(*!
<summary>Formats a failed typed predicate and reports it with the chain message.</summary>
<description>
Does not change operands or chain state. The receiver retains its first failure. Reporting exceptions
propagate to the enclosing test callback handler; an unprepared receiver is a configuration error.
</description>
<param name="expected">Typed expected operand used only for this diagnostic.</param>
<param name="expectation">Prefix identifying the failed predicate.</param>
*)
METHOD PRIVATE failComparison
VAR_INPUT
	expected : SINT;
	expectation : WSTRING(40);
END_VAR
VAR
	actualText : WSTRING(255);
	expectedText : WSTRING(255);
	diagnostic : TOF_Core.ERROR_MESSAGE;
END_VAR
actualText := TO_WSTRING(_Actual);
expectedText := TO_WSTRING(expected);

diagnostic := TOF_Core.WideStrings.Concat255(
	expectation,
	expectedText,
	", but was: ",
	actualText
);

TestServices.ReportAssertionFailure(
	testCase := _TestCase,
	message := _Message,
	sourceClassName := ClassName,
	defaultMessage := diagnostic
);
END_METHOD

END_FUNCTION_BLOCK

// ---- Assertions/TypedContexts/IntAssertionContext.TcPOU
(*
SPDX-FileCopyrightText: © 2026 Oleksandr Tiutyk <trofimich@gmail.com>
SPDX-License-Identifier: MIT
License: https://opensource.org/license/mit
*)

(*!
<summary>Provides fluent assertions on a copied INT value.</summary>
<description>
Copies actual into persistent instance storage before the entry method returns; literals and expression
results therefore remain valid throughout the immediate chain. Owns no heap allocation or pointed-to resource.
The message prefixes every failure until the next preparation. Finish one chain before starting another on
the owning Assertions provider. Use only from the owning test callback on one task, without reentry.
Obtain this context from the owning provider; direct unprepared use is unsupported.
Expected arguments use the declared IEC type; ordinary compiler conversions happen before comparison.
This context does not depend on another assertion context.
Object metadata is available before preparation; inherited equality compares instance identity.
</description>
*)

{attribute 'no_explicit_call' := 'do not call this function block directly'}
FUNCTION_BLOCK IntAssertionContext EXTENDS TOF_Core.Object
VAR_STAT
	{attribute 'hide'}
	_ClassName : STRING := __POUNAME();
END_VAR
VAR
	_Actual : INT;
	_TestCase : ITestCase;
	_Message : WSTRING(255);
END_VAR

(*!
<summary>Provides the implementation class name.</summary>
<description>
Borrowed read-only reference to compiler-initialized storage, valid throughout the instance lifetime.
Do not modify the returned reference; no ownership is transferred.
</description>
*)
{attribute 'monitoring' := 'call'}
PROPERTY ClassName : REFERENCE TO STRING
GET
ClassName REF= _ClassName;
END_GET
END_PROPERTY

(*!
<summary>Asserts that the actual value is strictly greater than expected.</summary>
<description>
Records failure without interrupting the callback; preserves the message for the rest of the chain.
</description>
<param name="expected">Expected value converted by the compiler to INT.</param>
*)
METHOD FINAL IsGreaterThan : REFERENCE TO IntAssertionContext
VAR_INPUT
	expected : INT;
END_VAR
IF _Actual <= expected THEN
	failComparison(
		expected := expected,
		expectation := "Expected value > "
	);
END_IF

IsGreaterThan REF= THIS^;
END_METHOD

(*!
<summary>Asserts that the actual value meets the inclusive lower boundary.</summary>
<description>
Records failure without interrupting the callback; preserves the message for the rest of the chain.
</description>
<param name="expected">Expected value converted by the compiler to INT.</param>
*)
METHOD FINAL IsGreaterThanOrEquals : REFERENCE TO IntAssertionContext
VAR_INPUT
	expected : INT;
END_VAR
IF _Actual < expected THEN
	failComparison(
		expected := expected,
		expectation := "Expected value >= "
	);
END_IF

IsGreaterThanOrEquals REF= THIS^;
END_METHOD

(*!
<summary>Asserts that the actual value is strictly less than expected.</summary>
<description>
Records failure without interrupting the callback; preserves the message for the rest of the chain.
</description>
<param name="expected">Expected value converted by the compiler to INT.</param>
*)
METHOD FINAL IsLessThan : REFERENCE TO IntAssertionContext
VAR_INPUT
	expected : INT;
END_VAR
IF _Actual >= expected THEN
	failComparison(
		expected := expected,
		expectation := "Expected value < "
	);
END_IF

IsLessThan REF= THIS^;
END_METHOD

(*!
<summary>Asserts that the actual value meets the inclusive upper boundary.</summary>
<description>
Records failure without interrupting the callback; preserves the message for the rest of the chain.
</description>
<param name="expected">Expected value converted by the compiler to INT.</param>
*)
METHOD FINAL IsLessThanOrEquals : REFERENCE TO IntAssertionContext
VAR_INPUT
	expected : INT;
END_VAR
IF _Actual > expected THEN
	failComparison(
		expected := expected,
		expectation := "Expected value <= "
	);
END_IF

IsLessThanOrEquals REF= THIS^;
END_METHOD

(*!
<summary>Provides the library namespace.</summary>
<description>
Borrowed read-only reference to the compiler-initialized namespace, valid throughout the instance lifetime.
Do not modify the returned reference; no ownership is transferred.
</description>
*)
{attribute 'monitoring' := 'call'}
PROPERTY NamespaceName : REFERENCE TO STRING
GET
NamespaceName REF= CurrentNamespace.Name;
END_GET
END_PROPERTY

(*!
<summary>Asserts inequality with the expected value.</summary>
<description>
Records failure without interrupting the callback; preserves the message for the rest of the chain.
</description>
<param name="expected">Expected value converted by the compiler to INT.</param>
*)
METHOD FINAL NotToBe : REFERENCE TO IntAssertionContext
VAR_INPUT
	expected : INT;
END_VAR
IF _Actual = expected THEN
	failComparison(
		expected := expected,
		expectation := "Expected value not to be: "
	);
END_IF

NotToBe REF= THIS^;
END_METHOD

(*!
<summary>Copies the actual operand and replaces the chain-wide message.</summary>
<description>
Called by the owning Assertions provider after it verifies the running test case.
No pointer to this method's input storage is retained. The receiver is borrowed until the next preparation;
the owning provider keeps it alive throughout the immediate chain.
</description>
<param name="actual">Value copied into this context.</param>
<param name="testCase">Borrowed failure receiver for the immediate chain.</param>
<param name="message">Copied diagnostic prefix, including empty to clear the previous prefix.</param>
*)
METHOD INTERNAL FINAL Prepare
VAR_INPUT
	actual : INT;
	testCase : ITestCase;
	message : WSTRING(255);
END_VAR
_Actual := actual;
_TestCase := testCase;
_Message := message;
END_METHOD

(*!
<summary>Reports the byte size of this concrete instance.</summary>
<description>
Includes inline fields and nested instances, but excludes separately allocated payloads.
Obtaining the size does not transfer ownership or validate an arbitrary address.
</description>
*)
{attribute 'monitoring' := 'call'}
PROPERTY SelfSize : ULINT
GET
SelfSize := XSIZEOF(THIS^);
END_GET
END_PROPERTY

(*!
<summary>Asserts equality with the expected value.</summary>
<description>
Records failure without interrupting the callback; preserves the message for the rest of the chain.
</description>
<param name="expected">Expected value converted by the compiler to INT.</param>
*)
METHOD FINAL ToBe : REFERENCE TO IntAssertionContext
VAR_INPUT
	expected : INT;
END_VAR
IF _Actual <> expected THEN
	failComparison(
		expected := expected,
		expectation := "Expected: "
	);
END_IF

ToBe REF= THIS^;
END_METHOD

(*!
<summary>Formats a failed typed predicate and reports it with the chain message.</summary>
<description>
Does not change operands or chain state. The receiver retains its first failure. Reporting exceptions
propagate to the enclosing test callback handler; an unprepared receiver is a configuration error.
</description>
<param name="expected">Typed expected operand used only for this diagnostic.</param>
<param name="expectation">Prefix identifying the failed predicate.</param>
*)
METHOD PRIVATE failComparison
VAR_INPUT
	expected : INT;
	expectation : WSTRING(40);
END_VAR
VAR
	actualText : WSTRING(255);
	expectedText : WSTRING(255);
	diagnostic : TOF_Core.ERROR_MESSAGE;
END_VAR
actualText := TO_WSTRING(_Actual);
expectedText := TO_WSTRING(expected);

diagnostic := TOF_Core.WideStrings.Concat255(
	expectation,
	expectedText,
	", but was: ",
	actualText
);

TestServices.ReportAssertionFailure(
	testCase := _TestCase,
	message := _Message,
	sourceClassName := ClassName,
	defaultMessage := diagnostic
);
END_METHOD

END_FUNCTION_BLOCK

// ---- Assertions/TypedContexts/DIntAssertionContext.TcPOU
(*
SPDX-FileCopyrightText: © 2026 Oleksandr Tiutyk <trofimich@gmail.com>
SPDX-License-Identifier: MIT
License: https://opensource.org/license/mit
*)

(*!
<summary>Provides fluent assertions on a copied DINT value.</summary>
<description>
Copies actual into persistent instance storage before the entry method returns; literals and expression
results therefore remain valid throughout the immediate chain. Owns no heap allocation or pointed-to resource.
The message prefixes every failure until the next preparation. Finish one chain before starting another on
the owning Assertions provider. Use only from the owning test callback on one task, without reentry.
Obtain this context from the owning provider; direct unprepared use is unsupported.
Expected arguments use the declared IEC type; ordinary compiler conversions happen before comparison.
This context does not depend on another assertion context.
Object metadata is available before preparation; inherited equality compares instance identity.
</description>
*)

{attribute 'no_explicit_call' := 'do not call this function block directly'}
FUNCTION_BLOCK DIntAssertionContext EXTENDS TOF_Core.Object
VAR_STAT
	{attribute 'hide'}
	_ClassName : STRING := __POUNAME();
END_VAR
VAR
	_Actual : DINT;
	_TestCase : ITestCase;
	_Message : WSTRING(255);
END_VAR

(*!
<summary>Provides the implementation class name.</summary>
<description>
Borrowed read-only reference to compiler-initialized storage, valid throughout the instance lifetime.
Do not modify the returned reference; no ownership is transferred.
</description>
*)
{attribute 'monitoring' := 'call'}
PROPERTY ClassName : REFERENCE TO STRING
GET
ClassName REF= _ClassName;
END_GET
END_PROPERTY

(*!
<summary>Asserts that the actual value is strictly greater than expected.</summary>
<description>
Records failure without interrupting the callback; preserves the message for the rest of the chain.
</description>
<param name="expected">Expected value converted by the compiler to DINT.</param>
*)
METHOD FINAL IsGreaterThan : REFERENCE TO DIntAssertionContext
VAR_INPUT
	expected : DINT;
END_VAR
IF _Actual <= expected THEN
	failComparison(
		expected := expected,
		expectation := "Expected value > "
	);
END_IF

IsGreaterThan REF= THIS^;
END_METHOD

(*!
<summary>Asserts that the actual value meets the inclusive lower boundary.</summary>
<description>
Records failure without interrupting the callback; preserves the message for the rest of the chain.
</description>
<param name="expected">Expected value converted by the compiler to DINT.</param>
*)
METHOD FINAL IsGreaterThanOrEquals : REFERENCE TO DIntAssertionContext
VAR_INPUT
	expected : DINT;
END_VAR
IF _Actual < expected THEN
	failComparison(
		expected := expected,
		expectation := "Expected value >= "
	);
END_IF

IsGreaterThanOrEquals REF= THIS^;
END_METHOD

(*!
<summary>Asserts that the actual value is strictly less than expected.</summary>
<description>
Records failure without interrupting the callback; preserves the message for the rest of the chain.
</description>
<param name="expected">Expected value converted by the compiler to DINT.</param>
*)
METHOD FINAL IsLessThan : REFERENCE TO DIntAssertionContext
VAR_INPUT
	expected : DINT;
END_VAR
IF _Actual >= expected THEN
	failComparison(
		expected := expected,
		expectation := "Expected value < "
	);
END_IF

IsLessThan REF= THIS^;
END_METHOD

(*!
<summary>Asserts that the actual value meets the inclusive upper boundary.</summary>
<description>
Records failure without interrupting the callback; preserves the message for the rest of the chain.
</description>
<param name="expected">Expected value converted by the compiler to DINT.</param>
*)
METHOD FINAL IsLessThanOrEquals : REFERENCE TO DIntAssertionContext
VAR_INPUT
	expected : DINT;
END_VAR
IF _Actual > expected THEN
	failComparison(
		expected := expected,
		expectation := "Expected value <= "
	);
END_IF

IsLessThanOrEquals REF= THIS^;
END_METHOD

(*!
<summary>Provides the library namespace.</summary>
<description>
Borrowed read-only reference to the compiler-initialized namespace, valid throughout the instance lifetime.
Do not modify the returned reference; no ownership is transferred.
</description>
*)
{attribute 'monitoring' := 'call'}
PROPERTY NamespaceName : REFERENCE TO STRING
GET
NamespaceName REF= CurrentNamespace.Name;
END_GET
END_PROPERTY

(*!
<summary>Asserts inequality with the expected value.</summary>
<description>
Records failure without interrupting the callback; preserves the message for the rest of the chain.
</description>
<param name="expected">Expected value converted by the compiler to DINT.</param>
*)
METHOD FINAL NotToBe : REFERENCE TO DIntAssertionContext
VAR_INPUT
	expected : DINT;
END_VAR
IF _Actual = expected THEN
	failComparison(
		expected := expected,
		expectation := "Expected value not to be: "
	);
END_IF

NotToBe REF= THIS^;
END_METHOD

(*!
<summary>Copies the actual operand and replaces the chain-wide message.</summary>
<description>
Called by the owning Assertions provider after it verifies the running test case.
No pointer to this method's input storage is retained. The receiver is borrowed until the next preparation;
the owning provider keeps it alive throughout the immediate chain.
</description>
<param name="actual">Value copied into this context.</param>
<param name="testCase">Borrowed failure receiver for the immediate chain.</param>
<param name="message">Copied diagnostic prefix, including empty to clear the previous prefix.</param>
*)
METHOD INTERNAL FINAL Prepare
VAR_INPUT
	actual : DINT;
	testCase : ITestCase;
	message : WSTRING(255);
END_VAR
_Actual := actual;
_TestCase := testCase;
_Message := message;
END_METHOD

(*!
<summary>Reports the byte size of this concrete instance.</summary>
<description>
Includes inline fields and nested instances, but excludes separately allocated payloads.
Obtaining the size does not transfer ownership or validate an arbitrary address.
</description>
*)
{attribute 'monitoring' := 'call'}
PROPERTY SelfSize : ULINT
GET
SelfSize := XSIZEOF(THIS^);
END_GET
END_PROPERTY

(*!
<summary>Asserts equality with the expected value.</summary>
<description>
Records failure without interrupting the callback; preserves the message for the rest of the chain.
</description>
<param name="expected">Expected value converted by the compiler to DINT.</param>
*)
METHOD FINAL ToBe : REFERENCE TO DIntAssertionContext
VAR_INPUT
	expected : DINT;
END_VAR
IF _Actual <> expected THEN
	failComparison(
		expected := expected,
		expectation := "Expected: "
	);
END_IF

ToBe REF= THIS^;
END_METHOD

(*!
<summary>Formats a failed typed predicate and reports it with the chain message.</summary>
<description>
Does not change operands or chain state. The receiver retains its first failure. Reporting exceptions
propagate to the enclosing test callback handler; an unprepared receiver is a configuration error.
</description>
<param name="expected">Typed expected operand used only for this diagnostic.</param>
<param name="expectation">Prefix identifying the failed predicate.</param>
*)
METHOD PRIVATE failComparison
VAR_INPUT
	expected : DINT;
	expectation : WSTRING(40);
END_VAR
VAR
	actualText : WSTRING(255);
	expectedText : WSTRING(255);
	diagnostic : TOF_Core.ERROR_MESSAGE;
END_VAR
actualText := TO_WSTRING(_Actual);
expectedText := TO_WSTRING(expected);

diagnostic := TOF_Core.WideStrings.Concat255(
	expectation,
	expectedText,
	", but was: ",
	actualText
);

TestServices.ReportAssertionFailure(
	testCase := _TestCase,
	message := _Message,
	sourceClassName := ClassName,
	defaultMessage := diagnostic
);
END_METHOD

END_FUNCTION_BLOCK

// ---- Assertions/TypedContexts/LIntAssertionContext.TcPOU
(*
SPDX-FileCopyrightText: © 2026 Oleksandr Tiutyk <trofimich@gmail.com>
SPDX-License-Identifier: MIT
License: https://opensource.org/license/mit
*)

(*!
<summary>Provides fluent assertions on a copied LINT value.</summary>
<description>
Copies actual into persistent instance storage before the entry method returns; literals and expression
results therefore remain valid throughout the immediate chain. Owns no heap allocation or pointed-to resource.
The message prefixes every failure until the next preparation. Finish one chain before starting another on
the owning Assertions provider. Use only from the owning test callback on one task, without reentry.
Obtain this context from the owning provider; direct unprepared use is unsupported.
Expected arguments use the declared IEC type; ordinary compiler conversions happen before comparison.
This context does not depend on another assertion context.
Object metadata is available before preparation; inherited equality compares instance identity.
</description>
*)

{attribute 'no_explicit_call' := 'do not call this function block directly'}
FUNCTION_BLOCK LIntAssertionContext EXTENDS TOF_Core.Object
VAR_STAT
	{attribute 'hide'}
	_ClassName : STRING := __POUNAME();
END_VAR
VAR
	_Actual : LINT;
	_TestCase : ITestCase;
	_Message : WSTRING(255);
END_VAR

(*!
<summary>Provides the implementation class name.</summary>
<description>
Borrowed read-only reference to compiler-initialized storage, valid throughout the instance lifetime.
Do not modify the returned reference; no ownership is transferred.
</description>
*)
{attribute 'monitoring' := 'call'}
PROPERTY ClassName : REFERENCE TO STRING
GET
ClassName REF= _ClassName;
END_GET
END_PROPERTY

(*!
<summary>Asserts that the actual value is strictly greater than expected.</summary>
<description>
Records failure without interrupting the callback; preserves the message for the rest of the chain.
</description>
<param name="expected">Expected value converted by the compiler to LINT.</param>
*)
METHOD FINAL IsGreaterThan : REFERENCE TO LIntAssertionContext
VAR_INPUT
	expected : LINT;
END_VAR
IF _Actual <= expected THEN
	failComparison(
		expected := expected,
		expectation := "Expected value > "
	);
END_IF

IsGreaterThan REF= THIS^;
END_METHOD

(*!
<summary>Asserts that the actual value meets the inclusive lower boundary.</summary>
<description>
Records failure without interrupting the callback; preserves the message for the rest of the chain.
</description>
<param name="expected">Expected value converted by the compiler to LINT.</param>
*)
METHOD FINAL IsGreaterThanOrEquals : REFERENCE TO LIntAssertionContext
VAR_INPUT
	expected : LINT;
END_VAR
IF _Actual < expected THEN
	failComparison(
		expected := expected,
		expectation := "Expected value >= "
	);
END_IF

IsGreaterThanOrEquals REF= THIS^;
END_METHOD

(*!
<summary>Asserts that the actual value is strictly less than expected.</summary>
<description>
Records failure without interrupting the callback; preserves the message for the rest of the chain.
</description>
<param name="expected">Expected value converted by the compiler to LINT.</param>
*)
METHOD FINAL IsLessThan : REFERENCE TO LIntAssertionContext
VAR_INPUT
	expected : LINT;
END_VAR
IF _Actual >= expected THEN
	failComparison(
		expected := expected,
		expectation := "Expected value < "
	);
END_IF

IsLessThan REF= THIS^;
END_METHOD

(*!
<summary>Asserts that the actual value meets the inclusive upper boundary.</summary>
<description>
Records failure without interrupting the callback; preserves the message for the rest of the chain.
</description>
<param name="expected">Expected value converted by the compiler to LINT.</param>
*)
METHOD FINAL IsLessThanOrEquals : REFERENCE TO LIntAssertionContext
VAR_INPUT
	expected : LINT;
END_VAR
IF _Actual > expected THEN
	failComparison(
		expected := expected,
		expectation := "Expected value <= "
	);
END_IF

IsLessThanOrEquals REF= THIS^;
END_METHOD

(*!
<summary>Provides the library namespace.</summary>
<description>
Borrowed read-only reference to the compiler-initialized namespace, valid throughout the instance lifetime.
Do not modify the returned reference; no ownership is transferred.
</description>
*)
{attribute 'monitoring' := 'call'}
PROPERTY NamespaceName : REFERENCE TO STRING
GET
NamespaceName REF= CurrentNamespace.Name;
END_GET
END_PROPERTY

(*!
<summary>Asserts inequality with the expected value.</summary>
<description>
Records failure without interrupting the callback; preserves the message for the rest of the chain.
</description>
<param name="expected">Expected value converted by the compiler to LINT.</param>
*)
METHOD FINAL NotToBe : REFERENCE TO LIntAssertionContext
VAR_INPUT
	expected : LINT;
END_VAR
IF _Actual = expected THEN
	failComparison(
		expected := expected,
		expectation := "Expected value not to be: "
	);
END_IF

NotToBe REF= THIS^;
END_METHOD

(*!
<summary>Copies the actual operand and replaces the chain-wide message.</summary>
<description>
Called by the owning Assertions provider after it verifies the running test case.
No pointer to this method's input storage is retained. The receiver is borrowed until the next preparation;
the owning provider keeps it alive throughout the immediate chain.
</description>
<param name="actual">Value copied into this context.</param>
<param name="testCase">Borrowed failure receiver for the immediate chain.</param>
<param name="message">Copied diagnostic prefix, including empty to clear the previous prefix.</param>
*)
METHOD INTERNAL FINAL Prepare
VAR_INPUT
	actual : LINT;
	testCase : ITestCase;
	message : WSTRING(255);
END_VAR
_Actual := actual;
_TestCase := testCase;
_Message := message;
END_METHOD

(*!
<summary>Reports the byte size of this concrete instance.</summary>
<description>
Includes inline fields and nested instances, but excludes separately allocated payloads.
Obtaining the size does not transfer ownership or validate an arbitrary address.
</description>
*)
{attribute 'monitoring' := 'call'}
PROPERTY SelfSize : ULINT
GET
SelfSize := XSIZEOF(THIS^);
END_GET
END_PROPERTY

(*!
<summary>Asserts equality with the expected value.</summary>
<description>
Records failure without interrupting the callback; preserves the message for the rest of the chain.
</description>
<param name="expected">Expected value converted by the compiler to LINT.</param>
*)
METHOD FINAL ToBe : REFERENCE TO LIntAssertionContext
VAR_INPUT
	expected : LINT;
END_VAR
IF _Actual <> expected THEN
	failComparison(
		expected := expected,
		expectation := "Expected: "
	);
END_IF

ToBe REF= THIS^;
END_METHOD

(*!
<summary>Formats a failed typed predicate and reports it with the chain message.</summary>
<description>
Does not change operands or chain state. The receiver retains its first failure. Reporting exceptions
propagate to the enclosing test callback handler; an unprepared receiver is a configuration error.
</description>
<param name="expected">Typed expected operand used only for this diagnostic.</param>
<param name="expectation">Prefix identifying the failed predicate.</param>
*)
METHOD PRIVATE failComparison
VAR_INPUT
	expected : LINT;
	expectation : WSTRING(40);
END_VAR
VAR
	actualText : WSTRING(255);
	expectedText : WSTRING(255);
	diagnostic : TOF_Core.ERROR_MESSAGE;
END_VAR
actualText := TO_WSTRING(_Actual);
expectedText := TO_WSTRING(expected);

diagnostic := TOF_Core.WideStrings.Concat255(
	expectation,
	expectedText,
	", but was: ",
	actualText
);

TestServices.ReportAssertionFailure(
	testCase := _TestCase,
	message := _Message,
	sourceClassName := ClassName,
	defaultMessage := diagnostic
);
END_METHOD

END_FUNCTION_BLOCK

// ---- Assertions/TypedContexts/USIntAssertionContext.TcPOU
(*
SPDX-FileCopyrightText: © 2026 Oleksandr Tiutyk <trofimich@gmail.com>
SPDX-License-Identifier: MIT
License: https://opensource.org/license/mit
*)

(*!
<summary>Provides fluent assertions on a copied USINT value.</summary>
<description>
Copies actual into persistent instance storage before the entry method returns; literals and expression
results therefore remain valid throughout the immediate chain. Owns no heap allocation or pointed-to resource.
The message prefixes every failure until the next preparation. Finish one chain before starting another on
the owning Assertions provider. Use only from the owning test callback on one task, without reentry.
Obtain this context from the owning provider; direct unprepared use is unsupported.
Expected arguments use the declared IEC type; ordinary compiler conversions happen before comparison.
This context does not depend on another assertion context.
Object metadata is available before preparation; inherited equality compares instance identity.
</description>
*)

{attribute 'no_explicit_call' := 'do not call this function block directly'}
FUNCTION_BLOCK USIntAssertionContext EXTENDS TOF_Core.Object
VAR_STAT
	{attribute 'hide'}
	_ClassName : STRING := __POUNAME();
END_VAR
VAR
	_Actual : USINT;
	_TestCase : ITestCase;
	_Message : WSTRING(255);
END_VAR

(*!
<summary>Provides the implementation class name.</summary>
<description>
Borrowed read-only reference to compiler-initialized storage, valid throughout the instance lifetime.
Do not modify the returned reference; no ownership is transferred.
</description>
*)
{attribute 'monitoring' := 'call'}
PROPERTY ClassName : REFERENCE TO STRING
GET
ClassName REF= _ClassName;
END_GET
END_PROPERTY

(*!
<summary>Asserts that the actual value is strictly greater than expected.</summary>
<description>
Records failure without interrupting the callback; preserves the message for the rest of the chain.
</description>
<param name="expected">Expected value converted by the compiler to USINT.</param>
*)
METHOD FINAL IsGreaterThan : REFERENCE TO USIntAssertionContext
VAR_INPUT
	expected : USINT;
END_VAR
IF _Actual <= expected THEN
	failComparison(
		expected := expected,
		expectation := "Expected value > "
	);
END_IF

IsGreaterThan REF= THIS^;
END_METHOD

(*!
<summary>Asserts that the actual value meets the inclusive lower boundary.</summary>
<description>
Records failure without interrupting the callback; preserves the message for the rest of the chain.
</description>
<param name="expected">Expected value converted by the compiler to USINT.</param>
*)
METHOD FINAL IsGreaterThanOrEquals : REFERENCE TO USIntAssertionContext
VAR_INPUT
	expected : USINT;
END_VAR
IF _Actual < expected THEN
	failComparison(
		expected := expected,
		expectation := "Expected value >= "
	);
END_IF

IsGreaterThanOrEquals REF= THIS^;
END_METHOD

(*!
<summary>Asserts that the actual value is strictly less than expected.</summary>
<description>
Records failure without interrupting the callback; preserves the message for the rest of the chain.
</description>
<param name="expected">Expected value converted by the compiler to USINT.</param>
*)
METHOD FINAL IsLessThan : REFERENCE TO USIntAssertionContext
VAR_INPUT
	expected : USINT;
END_VAR
IF _Actual >= expected THEN
	failComparison(
		expected := expected,
		expectation := "Expected value < "
	);
END_IF

IsLessThan REF= THIS^;
END_METHOD

(*!
<summary>Asserts that the actual value meets the inclusive upper boundary.</summary>
<description>
Records failure without interrupting the callback; preserves the message for the rest of the chain.
</description>
<param name="expected">Expected value converted by the compiler to USINT.</param>
*)
METHOD FINAL IsLessThanOrEquals : REFERENCE TO USIntAssertionContext
VAR_INPUT
	expected : USINT;
END_VAR
IF _Actual > expected THEN
	failComparison(
		expected := expected,
		expectation := "Expected value <= "
	);
END_IF

IsLessThanOrEquals REF= THIS^;
END_METHOD

(*!
<summary>Provides the library namespace.</summary>
<description>
Borrowed read-only reference to the compiler-initialized namespace, valid throughout the instance lifetime.
Do not modify the returned reference; no ownership is transferred.
</description>
*)
{attribute 'monitoring' := 'call'}
PROPERTY NamespaceName : REFERENCE TO STRING
GET
NamespaceName REF= CurrentNamespace.Name;
END_GET
END_PROPERTY

(*!
<summary>Asserts inequality with the expected value.</summary>
<description>
Records failure without interrupting the callback; preserves the message for the rest of the chain.
</description>
<param name="expected">Expected value converted by the compiler to USINT.</param>
*)
METHOD FINAL NotToBe : REFERENCE TO USIntAssertionContext
VAR_INPUT
	expected : USINT;
END_VAR
IF _Actual = expected THEN
	failComparison(
		expected := expected,
		expectation := "Expected value not to be: "
	);
END_IF

NotToBe REF= THIS^;
END_METHOD

(*!
<summary>Copies the actual operand and replaces the chain-wide message.</summary>
<description>
Called by the owning Assertions provider after it verifies the running test case.
No pointer to this method's input storage is retained. The receiver is borrowed until the next preparation;
the owning provider keeps it alive throughout the immediate chain.
</description>
<param name="actual">Value copied into this context.</param>
<param name="testCase">Borrowed failure receiver for the immediate chain.</param>
<param name="message">Copied diagnostic prefix, including empty to clear the previous prefix.</param>
*)
METHOD INTERNAL FINAL Prepare
VAR_INPUT
	actual : USINT;
	testCase : ITestCase;
	message : WSTRING(255);
END_VAR
_Actual := actual;
_TestCase := testCase;
_Message := message;
END_METHOD

(*!
<summary>Reports the byte size of this concrete instance.</summary>
<description>
Includes inline fields and nested instances, but excludes separately allocated payloads.
Obtaining the size does not transfer ownership or validate an arbitrary address.
</description>
*)
{attribute 'monitoring' := 'call'}
PROPERTY SelfSize : ULINT
GET
SelfSize := XSIZEOF(THIS^);
END_GET
END_PROPERTY

(*!
<summary>Asserts equality with the expected value.</summary>
<description>
Records failure without interrupting the callback; preserves the message for the rest of the chain.
</description>
<param name="expected">Expected value converted by the compiler to USINT.</param>
*)
METHOD FINAL ToBe : REFERENCE TO USIntAssertionContext
VAR_INPUT
	expected : USINT;
END_VAR
IF _Actual <> expected THEN
	failComparison(
		expected := expected,
		expectation := "Expected: "
	);
END_IF

ToBe REF= THIS^;
END_METHOD

(*!
<summary>Formats a failed typed predicate and reports it with the chain message.</summary>
<description>
Does not change operands or chain state. The receiver retains its first failure. Reporting exceptions
propagate to the enclosing test callback handler; an unprepared receiver is a configuration error.
</description>
<param name="expected">Typed expected operand used only for this diagnostic.</param>
<param name="expectation">Prefix identifying the failed predicate.</param>
*)
METHOD PRIVATE failComparison
VAR_INPUT
	expected : USINT;
	expectation : WSTRING(40);
END_VAR
VAR
	actualText : WSTRING(255);
	expectedText : WSTRING(255);
	diagnostic : TOF_Core.ERROR_MESSAGE;
END_VAR
actualText := TO_WSTRING(_Actual);
expectedText := TO_WSTRING(expected);

diagnostic := TOF_Core.WideStrings.Concat255(
	expectation,
	expectedText,
	", but was: ",
	actualText
);

TestServices.ReportAssertionFailure(
	testCase := _TestCase,
	message := _Message,
	sourceClassName := ClassName,
	defaultMessage := diagnostic
);
END_METHOD

END_FUNCTION_BLOCK

// ---- Assertions/TypedContexts/UIntAssertionContext.TcPOU
(*
SPDX-FileCopyrightText: © 2026 Oleksandr Tiutyk <trofimich@gmail.com>
SPDX-License-Identifier: MIT
License: https://opensource.org/license/mit
*)

(*!
<summary>Provides fluent assertions on a copied UINT value.</summary>
<description>
Copies actual into persistent instance storage before the entry method returns; literals and expression
results therefore remain valid throughout the immediate chain. Owns no heap allocation or pointed-to resource.
The message prefixes every failure until the next preparation. Finish one chain before starting another on
the owning Assertions provider. Use only from the owning test callback on one task, without reentry.
Obtain this context from the owning provider; direct unprepared use is unsupported.
Expected arguments use the declared IEC type; ordinary compiler conversions happen before comparison.
This context does not depend on another assertion context.
Object metadata is available before preparation; inherited equality compares instance identity.
</description>
*)

{attribute 'no_explicit_call' := 'do not call this function block directly'}
FUNCTION_BLOCK UIntAssertionContext EXTENDS TOF_Core.Object
VAR_STAT
	{attribute 'hide'}
	_ClassName : STRING := __POUNAME();
END_VAR
VAR
	_Actual : UINT;
	_TestCase : ITestCase;
	_Message : WSTRING(255);
END_VAR

(*!
<summary>Provides the implementation class name.</summary>
<description>
Borrowed read-only reference to compiler-initialized storage, valid throughout the instance lifetime.
Do not modify the returned reference; no ownership is transferred.
</description>
*)
{attribute 'monitoring' := 'call'}
PROPERTY ClassName : REFERENCE TO STRING
GET
ClassName REF= _ClassName;
END_GET
END_PROPERTY

(*!
<summary>Asserts that the actual value is strictly greater than expected.</summary>
<description>
Records failure without interrupting the callback; preserves the message for the rest of the chain.
</description>
<param name="expected">Expected value converted by the compiler to UINT.</param>
*)
METHOD FINAL IsGreaterThan : REFERENCE TO UIntAssertionContext
VAR_INPUT
	expected : UINT;
END_VAR
IF _Actual <= expected THEN
	failComparison(
		expected := expected,
		expectation := "Expected value > "
	);
END_IF

IsGreaterThan REF= THIS^;
END_METHOD

(*!
<summary>Asserts that the actual value meets the inclusive lower boundary.</summary>
<description>
Records failure without interrupting the callback; preserves the message for the rest of the chain.
</description>
<param name="expected">Expected value converted by the compiler to UINT.</param>
*)
METHOD FINAL IsGreaterThanOrEquals : REFERENCE TO UIntAssertionContext
VAR_INPUT
	expected : UINT;
END_VAR
IF _Actual < expected THEN
	failComparison(
		expected := expected,
		expectation := "Expected value >= "
	);
END_IF

IsGreaterThanOrEquals REF= THIS^;
END_METHOD

(*!
<summary>Asserts that the actual value is strictly less than expected.</summary>
<description>
Records failure without interrupting the callback; preserves the message for the rest of the chain.
</description>
<param name="expected">Expected value converted by the compiler to UINT.</param>
*)
METHOD FINAL IsLessThan : REFERENCE TO UIntAssertionContext
VAR_INPUT
	expected : UINT;
END_VAR
IF _Actual >= expected THEN
	failComparison(
		expected := expected,
		expectation := "Expected value < "
	);
END_IF

IsLessThan REF= THIS^;
END_METHOD

(*!
<summary>Asserts that the actual value meets the inclusive upper boundary.</summary>
<description>
Records failure without interrupting the callback; preserves the message for the rest of the chain.
</description>
<param name="expected">Expected value converted by the compiler to UINT.</param>
*)
METHOD FINAL IsLessThanOrEquals : REFERENCE TO UIntAssertionContext
VAR_INPUT
	expected : UINT;
END_VAR
IF _Actual > expected THEN
	failComparison(
		expected := expected,
		expectation := "Expected value <= "
	);
END_IF

IsLessThanOrEquals REF= THIS^;
END_METHOD

(*!
<summary>Provides the library namespace.</summary>
<description>
Borrowed read-only reference to the compiler-initialized namespace, valid throughout the instance lifetime.
Do not modify the returned reference; no ownership is transferred.
</description>
*)
{attribute 'monitoring' := 'call'}
PROPERTY NamespaceName : REFERENCE TO STRING
GET
NamespaceName REF= CurrentNamespace.Name;
END_GET
END_PROPERTY

(*!
<summary>Asserts inequality with the expected value.</summary>
<description>
Records failure without interrupting the callback; preserves the message for the rest of the chain.
</description>
<param name="expected">Expected value converted by the compiler to UINT.</param>
*)
METHOD FINAL NotToBe : REFERENCE TO UIntAssertionContext
VAR_INPUT
	expected : UINT;
END_VAR
IF _Actual = expected THEN
	failComparison(
		expected := expected,
		expectation := "Expected value not to be: "
	);
END_IF

NotToBe REF= THIS^;
END_METHOD

(*!
<summary>Copies the actual operand and replaces the chain-wide message.</summary>
<description>
Called by the owning Assertions provider after it verifies the running test case.
No pointer to this method's input storage is retained. The receiver is borrowed until the next preparation;
the owning provider keeps it alive throughout the immediate chain.
</description>
<param name="actual">Value copied into this context.</param>
<param name="testCase">Borrowed failure receiver for the immediate chain.</param>
<param name="message">Copied diagnostic prefix, including empty to clear the previous prefix.</param>
*)
METHOD INTERNAL FINAL Prepare
VAR_INPUT
	actual : UINT;
	testCase : ITestCase;
	message : WSTRING(255);
END_VAR
_Actual := actual;
_TestCase := testCase;
_Message := message;
END_METHOD

(*!
<summary>Reports the byte size of this concrete instance.</summary>
<description>
Includes inline fields and nested instances, but excludes separately allocated payloads.
Obtaining the size does not transfer ownership or validate an arbitrary address.
</description>
*)
{attribute 'monitoring' := 'call'}
PROPERTY SelfSize : ULINT
GET
SelfSize := XSIZEOF(THIS^);
END_GET
END_PROPERTY

(*!
<summary>Asserts equality with the expected value.</summary>
<description>
Records failure without interrupting the callback; preserves the message for the rest of the chain.
</description>
<param name="expected">Expected value converted by the compiler to UINT.</param>
*)
METHOD FINAL ToBe : REFERENCE TO UIntAssertionContext
VAR_INPUT
	expected : UINT;
END_VAR
IF _Actual <> expected THEN
	failComparison(
		expected := expected,
		expectation := "Expected: "
	);
END_IF

ToBe REF= THIS^;
END_METHOD

(*!
<summary>Formats a failed typed predicate and reports it with the chain message.</summary>
<description>
Does not change operands or chain state. The receiver retains its first failure. Reporting exceptions
propagate to the enclosing test callback handler; an unprepared receiver is a configuration error.
</description>
<param name="expected">Typed expected operand used only for this diagnostic.</param>
<param name="expectation">Prefix identifying the failed predicate.</param>
*)
METHOD PRIVATE failComparison
VAR_INPUT
	expected : UINT;
	expectation : WSTRING(40);
END_VAR
VAR
	actualText : WSTRING(255);
	expectedText : WSTRING(255);
	diagnostic : TOF_Core.ERROR_MESSAGE;
END_VAR
actualText := TO_WSTRING(_Actual);
expectedText := TO_WSTRING(expected);

diagnostic := TOF_Core.WideStrings.Concat255(
	expectation,
	expectedText,
	", but was: ",
	actualText
);

TestServices.ReportAssertionFailure(
	testCase := _TestCase,
	message := _Message,
	sourceClassName := ClassName,
	defaultMessage := diagnostic
);
END_METHOD

END_FUNCTION_BLOCK

// ---- Assertions/TypedContexts/UDIntAssertionContext.TcPOU
(*
SPDX-FileCopyrightText: © 2026 Oleksandr Tiutyk <trofimich@gmail.com>
SPDX-License-Identifier: MIT
License: https://opensource.org/license/mit
*)

(*!
<summary>Provides fluent assertions on a copied UDINT value.</summary>
<description>
Copies actual into persistent instance storage before the entry method returns; literals and expression
results therefore remain valid throughout the immediate chain. Owns no heap allocation or pointed-to resource.
The message prefixes every failure until the next preparation. Finish one chain before starting another on
the owning Assertions provider. Use only from the owning test callback on one task, without reentry.
Obtain this context from the owning provider; direct unprepared use is unsupported.
Expected arguments use the declared IEC type; ordinary compiler conversions happen before comparison.
This context does not depend on another assertion context.
Object metadata is available before preparation; inherited equality compares instance identity.
</description>
*)

{attribute 'no_explicit_call' := 'do not call this function block directly'}
FUNCTION_BLOCK UDIntAssertionContext EXTENDS TOF_Core.Object
VAR_STAT
	{attribute 'hide'}
	_ClassName : STRING := __POUNAME();
END_VAR
VAR
	_Actual : UDINT;
	_TestCase : ITestCase;
	_Message : WSTRING(255);
END_VAR

(*!
<summary>Provides the implementation class name.</summary>
<description>
Borrowed read-only reference to compiler-initialized storage, valid throughout the instance lifetime.
Do not modify the returned reference; no ownership is transferred.
</description>
*)
{attribute 'monitoring' := 'call'}
PROPERTY ClassName : REFERENCE TO STRING
GET
ClassName REF= _ClassName;
END_GET
END_PROPERTY

(*!
<summary>Asserts that the actual value is strictly greater than expected.</summary>
<description>
Records failure without interrupting the callback; preserves the message for the rest of the chain.
</description>
<param name="expected">Expected value converted by the compiler to UDINT.</param>
*)
METHOD FINAL IsGreaterThan : REFERENCE TO UDIntAssertionContext
VAR_INPUT
	expected : UDINT;
END_VAR
IF _Actual <= expected THEN
	failComparison(
		expected := expected,
		expectation := "Expected value > "
	);
END_IF

IsGreaterThan REF= THIS^;
END_METHOD

(*!
<summary>Asserts that the actual value meets the inclusive lower boundary.</summary>
<description>
Records failure without interrupting the callback; preserves the message for the rest of the chain.
</description>
<param name="expected">Expected value converted by the compiler to UDINT.</param>
*)
METHOD FINAL IsGreaterThanOrEquals : REFERENCE TO UDIntAssertionContext
VAR_INPUT
	expected : UDINT;
END_VAR
IF _Actual < expected THEN
	failComparison(
		expected := expected,
		expectation := "Expected value >= "
	);
END_IF

IsGreaterThanOrEquals REF= THIS^;
END_METHOD

(*!
<summary>Asserts that the actual value is strictly less than expected.</summary>
<description>
Records failure without interrupting the callback; preserves the message for the rest of the chain.
</description>
<param name="expected">Expected value converted by the compiler to UDINT.</param>
*)
METHOD FINAL IsLessThan : REFERENCE TO UDIntAssertionContext
VAR_INPUT
	expected : UDINT;
END_VAR
IF _Actual >= expected THEN
	failComparison(
		expected := expected,
		expectation := "Expected value < "
	);
END_IF

IsLessThan REF= THIS^;
END_METHOD

(*!
<summary>Asserts that the actual value meets the inclusive upper boundary.</summary>
<description>
Records failure without interrupting the callback; preserves the message for the rest of the chain.
</description>
<param name="expected">Expected value converted by the compiler to UDINT.</param>
*)
METHOD FINAL IsLessThanOrEquals : REFERENCE TO UDIntAssertionContext
VAR_INPUT
	expected : UDINT;
END_VAR
IF _Actual > expected THEN
	failComparison(
		expected := expected,
		expectation := "Expected value <= "
	);
END_IF

IsLessThanOrEquals REF= THIS^;
END_METHOD

(*!
<summary>Provides the library namespace.</summary>
<description>
Borrowed read-only reference to the compiler-initialized namespace, valid throughout the instance lifetime.
Do not modify the returned reference; no ownership is transferred.
</description>
*)
{attribute 'monitoring' := 'call'}
PROPERTY NamespaceName : REFERENCE TO STRING
GET
NamespaceName REF= CurrentNamespace.Name;
END_GET
END_PROPERTY

(*!
<summary>Asserts inequality with the expected value.</summary>
<description>
Records failure without interrupting the callback; preserves the message for the rest of the chain.
</description>
<param name="expected">Expected value converted by the compiler to UDINT.</param>
*)
METHOD FINAL NotToBe : REFERENCE TO UDIntAssertionContext
VAR_INPUT
	expected : UDINT;
END_VAR
IF _Actual = expected THEN
	failComparison(
		expected := expected,
		expectation := "Expected value not to be: "
	);
END_IF

NotToBe REF= THIS^;
END_METHOD

(*!
<summary>Copies the actual operand and replaces the chain-wide message.</summary>
<description>
Called by the owning Assertions provider after it verifies the running test case.
No pointer to this method's input storage is retained. The receiver is borrowed until the next preparation;
the owning provider keeps it alive throughout the immediate chain.
</description>
<param name="actual">Value copied into this context.</param>
<param name="testCase">Borrowed failure receiver for the immediate chain.</param>
<param name="message">Copied diagnostic prefix, including empty to clear the previous prefix.</param>
*)
METHOD INTERNAL FINAL Prepare
VAR_INPUT
	actual : UDINT;
	testCase : ITestCase;
	message : WSTRING(255);
END_VAR
_Actual := actual;
_TestCase := testCase;
_Message := message;
END_METHOD

(*!
<summary>Reports the byte size of this concrete instance.</summary>
<description>
Includes inline fields and nested instances, but excludes separately allocated payloads.
Obtaining the size does not transfer ownership or validate an arbitrary address.
</description>
*)
{attribute 'monitoring' := 'call'}
PROPERTY SelfSize : ULINT
GET
SelfSize := XSIZEOF(THIS^);
END_GET
END_PROPERTY

(*!
<summary>Asserts equality with the expected value.</summary>
<description>
Records failure without interrupting the callback; preserves the message for the rest of the chain.
</description>
<param name="expected">Expected value converted by the compiler to UDINT.</param>
*)
METHOD FINAL ToBe : REFERENCE TO UDIntAssertionContext
VAR_INPUT
	expected : UDINT;
END_VAR
IF _Actual <> expected THEN
	failComparison(
		expected := expected,
		expectation := "Expected: "
	);
END_IF

ToBe REF= THIS^;
END_METHOD

(*!
<summary>Formats a failed typed predicate and reports it with the chain message.</summary>
<description>
Does not change operands or chain state. The receiver retains its first failure. Reporting exceptions
propagate to the enclosing test callback handler; an unprepared receiver is a configuration error.
</description>
<param name="expected">Typed expected operand used only for this diagnostic.</param>
<param name="expectation">Prefix identifying the failed predicate.</param>
*)
METHOD PRIVATE failComparison
VAR_INPUT
	expected : UDINT;
	expectation : WSTRING(40);
END_VAR
VAR
	actualText : WSTRING(255);
	expectedText : WSTRING(255);
	diagnostic : TOF_Core.ERROR_MESSAGE;
END_VAR
actualText := TO_WSTRING(_Actual);
expectedText := TO_WSTRING(expected);

diagnostic := TOF_Core.WideStrings.Concat255(
	expectation,
	expectedText,
	", but was: ",
	actualText
);

TestServices.ReportAssertionFailure(
	testCase := _TestCase,
	message := _Message,
	sourceClassName := ClassName,
	defaultMessage := diagnostic
);
END_METHOD

END_FUNCTION_BLOCK

// ---- Assertions/TypedContexts/ULIntAssertionContext.TcPOU
(*
SPDX-FileCopyrightText: © 2026 Oleksandr Tiutyk <trofimich@gmail.com>
SPDX-License-Identifier: MIT
License: https://opensource.org/license/mit
*)

(*!
<summary>Provides fluent assertions on a copied ULINT value.</summary>
<description>
Copies actual into persistent instance storage before the entry method returns; literals and expression
results therefore remain valid throughout the immediate chain. Owns no heap allocation or pointed-to resource.
The message prefixes every failure until the next preparation. Finish one chain before starting another on
the owning Assertions provider. Use only from the owning test callback on one task, without reentry.
Obtain this context from the owning provider; direct unprepared use is unsupported.
Expected arguments use the declared IEC type; ordinary compiler conversions happen before comparison.
This context does not depend on another assertion context.
Object metadata is available before preparation; inherited equality compares instance identity.
</description>
*)

{attribute 'no_explicit_call' := 'do not call this function block directly'}
FUNCTION_BLOCK ULIntAssertionContext EXTENDS TOF_Core.Object
VAR_STAT
	{attribute 'hide'}
	_ClassName : STRING := __POUNAME();
END_VAR
VAR
	_Actual : ULINT;
	_TestCase : ITestCase;
	_Message : WSTRING(255);
END_VAR

(*!
<summary>Provides the implementation class name.</summary>
<description>
Borrowed read-only reference to compiler-initialized storage, valid throughout the instance lifetime.
Do not modify the returned reference; no ownership is transferred.
</description>
*)
{attribute 'monitoring' := 'call'}
PROPERTY ClassName : REFERENCE TO STRING
GET
ClassName REF= _ClassName;
END_GET
END_PROPERTY

(*!
<summary>Asserts that the actual value is strictly greater than expected.</summary>
<description>
Records failure without interrupting the callback; preserves the message for the rest of the chain.
</description>
<param name="expected">Expected value converted by the compiler to ULINT.</param>
*)
METHOD FINAL IsGreaterThan : REFERENCE TO ULIntAssertionContext
VAR_INPUT
	expected : ULINT;
END_VAR
IF _Actual <= expected THEN
	failComparison(
		expected := expected,
		expectation := "Expected value > "
	);
END_IF

IsGreaterThan REF= THIS^;
END_METHOD

(*!
<summary>Asserts that the actual value meets the inclusive lower boundary.</summary>
<description>
Records failure without interrupting the callback; preserves the message for the rest of the chain.
</description>
<param name="expected">Expected value converted by the compiler to ULINT.</param>
*)
METHOD FINAL IsGreaterThanOrEquals : REFERENCE TO ULIntAssertionContext
VAR_INPUT
	expected : ULINT;
END_VAR
IF _Actual < expected THEN
	failComparison(
		expected := expected,
		expectation := "Expected value >= "
	);
END_IF

IsGreaterThanOrEquals REF= THIS^;
END_METHOD

(*!
<summary>Asserts that the actual value is strictly less than expected.</summary>
<description>
Records failure without interrupting the callback; preserves the message for the rest of the chain.
</description>
<param name="expected">Expected value converted by the compiler to ULINT.</param>
*)
METHOD FINAL IsLessThan : REFERENCE TO ULIntAssertionContext
VAR_INPUT
	expected : ULINT;
END_VAR
IF _Actual >= expected THEN
	failComparison(
		expected := expected,
		expectation := "Expected value < "
	);
END_IF

IsLessThan REF= THIS^;
END_METHOD

(*!
<summary>Asserts that the actual value meets the inclusive upper boundary.</summary>
<description>
Records failure without interrupting the callback; preserves the message for the rest of the chain.
</description>
<param name="expected">Expected value converted by the compiler to ULINT.</param>
*)
METHOD FINAL IsLessThanOrEquals : REFERENCE TO ULIntAssertionContext
VAR_INPUT
	expected : ULINT;
END_VAR
IF _Actual > expected THEN
	failComparison(
		expected := expected,
		expectation := "Expected value <= "
	);
END_IF

IsLessThanOrEquals REF= THIS^;
END_METHOD

(*!
<summary>Provides the library namespace.</summary>
<description>
Borrowed read-only reference to the compiler-initialized namespace, valid throughout the instance lifetime.
Do not modify the returned reference; no ownership is transferred.
</description>
*)
{attribute 'monitoring' := 'call'}
PROPERTY NamespaceName : REFERENCE TO STRING
GET
NamespaceName REF= CurrentNamespace.Name;
END_GET
END_PROPERTY

(*!
<summary>Asserts inequality with the expected value.</summary>
<description>
Records failure without interrupting the callback; preserves the message for the rest of the chain.
</description>
<param name="expected">Expected value converted by the compiler to ULINT.</param>
*)
METHOD FINAL NotToBe : REFERENCE TO ULIntAssertionContext
VAR_INPUT
	expected : ULINT;
END_VAR
IF _Actual = expected THEN
	failComparison(
		expected := expected,
		expectation := "Expected value not to be: "
	);
END_IF

NotToBe REF= THIS^;
END_METHOD

(*!
<summary>Copies the actual operand and replaces the chain-wide message.</summary>
<description>
Called by the owning Assertions provider after it verifies the running test case.
No pointer to this method's input storage is retained. The receiver is borrowed until the next preparation;
the owning provider keeps it alive throughout the immediate chain.
</description>
<param name="actual">Value copied into this context.</param>
<param name="testCase">Borrowed failure receiver for the immediate chain.</param>
<param name="message">Copied diagnostic prefix, including empty to clear the previous prefix.</param>
*)
METHOD INTERNAL FINAL Prepare
VAR_INPUT
	actual : ULINT;
	testCase : ITestCase;
	message : WSTRING(255);
END_VAR
_Actual := actual;
_TestCase := testCase;
_Message := message;
END_METHOD

(*!
<summary>Reports the byte size of this concrete instance.</summary>
<description>
Includes inline fields and nested instances, but excludes separately allocated payloads.
Obtaining the size does not transfer ownership or validate an arbitrary address.
</description>
*)
{attribute 'monitoring' := 'call'}
PROPERTY SelfSize : ULINT
GET
SelfSize := XSIZEOF(THIS^);
END_GET
END_PROPERTY

(*!
<summary>Asserts equality with the expected value.</summary>
<description>
Records failure without interrupting the callback; preserves the message for the rest of the chain.
</description>
<param name="expected">Expected value converted by the compiler to ULINT.</param>
*)
METHOD FINAL ToBe : REFERENCE TO ULIntAssertionContext
VAR_INPUT
	expected : ULINT;
END_VAR
IF _Actual <> expected THEN
	failComparison(
		expected := expected,
		expectation := "Expected: "
	);
END_IF

ToBe REF= THIS^;
END_METHOD

(*!
<summary>Formats a failed typed predicate and reports it with the chain message.</summary>
<description>
Does not change operands or chain state. The receiver retains its first failure. Reporting exceptions
propagate to the enclosing test callback handler; an unprepared receiver is a configuration error.
</description>
<param name="expected">Typed expected operand used only for this diagnostic.</param>
<param name="expectation">Prefix identifying the failed predicate.</param>
*)
METHOD PRIVATE failComparison
VAR_INPUT
	expected : ULINT;
	expectation : WSTRING(40);
END_VAR
VAR
	actualText : WSTRING(255);
	expectedText : WSTRING(255);
	diagnostic : TOF_Core.ERROR_MESSAGE;
END_VAR
actualText := TO_WSTRING(_Actual);
expectedText := TO_WSTRING(expected);

diagnostic := TOF_Core.WideStrings.Concat255(
	expectation,
	expectedText,
	", but was: ",
	actualText
);

TestServices.ReportAssertionFailure(
	testCase := _TestCase,
	message := _Message,
	sourceClassName := ClassName,
	defaultMessage := diagnostic
);
END_METHOD

END_FUNCTION_BLOCK

// ---- Assertions/TypedContexts/ByteAssertionContext.TcPOU
(*
SPDX-FileCopyrightText: © 2026 Oleksandr Tiutyk <trofimich@gmail.com>
SPDX-License-Identifier: MIT
License: https://opensource.org/license/mit
*)

(*!
<summary>Provides fluent assertions on a copied BYTE value.</summary>
<description>
Copies actual into persistent instance storage before the entry method returns; literals and expression
results therefore remain valid throughout the immediate chain. Owns no heap allocation or pointed-to resource.
The message prefixes every failure until the next preparation. Finish one chain before starting another on
the owning Assertions provider. Use only from the owning test callback on one task, without reentry.
Obtain this context from the owning provider; direct unprepared use is unsupported.
Expected arguments use the declared IEC type; ordinary compiler conversions happen before comparison.
This context does not depend on another assertion context.
Object metadata is available before preparation; inherited equality compares instance identity.
</description>
*)

{attribute 'no_explicit_call' := 'do not call this function block directly'}
FUNCTION_BLOCK ByteAssertionContext EXTENDS TOF_Core.Object
VAR_STAT
	{attribute 'hide'}
	_ClassName : STRING := __POUNAME();
END_VAR
VAR
	_Actual : BYTE;
	_TestCase : ITestCase;
	_Message : WSTRING(255);
END_VAR

(*!
<summary>Provides the implementation class name.</summary>
<description>
Borrowed read-only reference to compiler-initialized storage, valid throughout the instance lifetime.
Do not modify the returned reference; no ownership is transferred.
</description>
*)
{attribute 'monitoring' := 'call'}
PROPERTY ClassName : REFERENCE TO STRING
GET
ClassName REF= _ClassName;
END_GET
END_PROPERTY

(*!
<summary>Asserts that the actual value is strictly greater than expected.</summary>
<description>
Records failure without interrupting the callback; preserves the message for the rest of the chain.
</description>
<param name="expected">Expected value converted by the compiler to BYTE.</param>
*)
METHOD FINAL IsGreaterThan : REFERENCE TO ByteAssertionContext
VAR_INPUT
	expected : BYTE;
END_VAR
IF _Actual <= expected THEN
	failComparison(
		expected := expected,
		expectation := "Expected value > "
	);
END_IF

IsGreaterThan REF= THIS^;
END_METHOD

(*!
<summary>Asserts that the actual value meets the inclusive lower boundary.</summary>
<description>
Records failure without interrupting the callback; preserves the message for the rest of the chain.
</description>
<param name="expected">Expected value converted by the compiler to BYTE.</param>
*)
METHOD FINAL IsGreaterThanOrEquals : REFERENCE TO ByteAssertionContext
VAR_INPUT
	expected : BYTE;
END_VAR
IF _Actual < expected THEN
	failComparison(
		expected := expected,
		expectation := "Expected value >= "
	);
END_IF

IsGreaterThanOrEquals REF= THIS^;
END_METHOD

(*!
<summary>Asserts that the actual value is strictly less than expected.</summary>
<description>
Records failure without interrupting the callback; preserves the message for the rest of the chain.
</description>
<param name="expected">Expected value converted by the compiler to BYTE.</param>
*)
METHOD FINAL IsLessThan : REFERENCE TO ByteAssertionContext
VAR_INPUT
	expected : BYTE;
END_VAR
IF _Actual >= expected THEN
	failComparison(
		expected := expected,
		expectation := "Expected value < "
	);
END_IF

IsLessThan REF= THIS^;
END_METHOD

(*!
<summary>Asserts that the actual value meets the inclusive upper boundary.</summary>
<description>
Records failure without interrupting the callback; preserves the message for the rest of the chain.
</description>
<param name="expected">Expected value converted by the compiler to BYTE.</param>
*)
METHOD FINAL IsLessThanOrEquals : REFERENCE TO ByteAssertionContext
VAR_INPUT
	expected : BYTE;
END_VAR
IF _Actual > expected THEN
	failComparison(
		expected := expected,
		expectation := "Expected value <= "
	);
END_IF

IsLessThanOrEquals REF= THIS^;
END_METHOD

(*!
<summary>Provides the library namespace.</summary>
<description>
Borrowed read-only reference to the compiler-initialized namespace, valid throughout the instance lifetime.
Do not modify the returned reference; no ownership is transferred.
</description>
*)
{attribute 'monitoring' := 'call'}
PROPERTY NamespaceName : REFERENCE TO STRING
GET
NamespaceName REF= CurrentNamespace.Name;
END_GET
END_PROPERTY

(*!
<summary>Asserts inequality with the expected value.</summary>
<description>
Records failure without interrupting the callback; preserves the message for the rest of the chain.
</description>
<param name="expected">Expected value converted by the compiler to BYTE.</param>
*)
METHOD FINAL NotToBe : REFERENCE TO ByteAssertionContext
VAR_INPUT
	expected : BYTE;
END_VAR
IF _Actual = expected THEN
	failComparison(
		expected := expected,
		expectation := "Expected value not to be: "
	);
END_IF

NotToBe REF= THIS^;
END_METHOD

(*!
<summary>Copies the actual operand and replaces the chain-wide message.</summary>
<description>
Called by the owning Assertions provider after it verifies the running test case.
No pointer to this method's input storage is retained. The receiver is borrowed until the next preparation;
the owning provider keeps it alive throughout the immediate chain.
</description>
<param name="actual">Value copied into this context.</param>
<param name="testCase">Borrowed failure receiver for the immediate chain.</param>
<param name="message">Copied diagnostic prefix, including empty to clear the previous prefix.</param>
*)
METHOD INTERNAL FINAL Prepare
VAR_INPUT
	actual : BYTE;
	testCase : ITestCase;
END_VAR
VAR_IN_OUT CONSTANT
	message : WSTRING(255);
END_VAR
_Actual := actual;
_TestCase := testCase;
_Message := message;
END_METHOD

(*!
<summary>Reports the byte size of this concrete instance.</summary>
<description>
Includes inline fields and nested instances, but excludes separately allocated payloads.
Obtaining the size does not transfer ownership or validate an arbitrary address.
</description>
*)
{attribute 'monitoring' := 'call'}
PROPERTY SelfSize : ULINT
GET
SelfSize := XSIZEOF(THIS^);
END_GET
END_PROPERTY

(*!
<summary>Asserts equality with the expected value.</summary>
<description>
Records failure without interrupting the callback; preserves the message for the rest of the chain.
</description>
<param name="expected">Expected value converted by the compiler to BYTE.</param>
*)
METHOD FINAL ToBe : REFERENCE TO ByteAssertionContext
VAR_INPUT
	expected : BYTE;
END_VAR
IF _Actual <> expected THEN
	failComparison(
		expected := expected,
		expectation := "Expected: "
	);
END_IF

ToBe REF= THIS^;
END_METHOD

(*!
<summary>Formats a failed typed predicate and reports it with the chain message.</summary>
<description>
Does not change operands or chain state. The receiver retains its first failure. Reporting exceptions
propagate to the enclosing test callback handler; an unprepared receiver is a configuration error.
</description>
<param name="expected">Typed expected operand used only for this diagnostic.</param>
<param name="expectation">Prefix identifying the failed predicate.</param>
*)
METHOD PRIVATE failComparison
VAR_INPUT
	expected : BYTE;
	expectation : WSTRING(40);
END_VAR
VAR
	actualText : WSTRING(255);
	expectedText : WSTRING(255);
	diagnostic : TOF_Core.ERROR_MESSAGE;
END_VAR
actualText := TO_WSTRING(TO_USINT(_Actual));
expectedText := TO_WSTRING(TO_USINT(expected));

diagnostic := TOF_Core.WideStrings.Concat255(
	expectation,
	expectedText,
	", but was: ",
	actualText
);

TestServices.ReportAssertionFailure(
	testCase := _TestCase,
	message := _Message,
	sourceClassName := ClassName,
	defaultMessage := diagnostic
);
END_METHOD

END_FUNCTION_BLOCK

// ---- Assertions/TypedContexts/WordAssertionContext.TcPOU
(*
SPDX-FileCopyrightText: © 2026 Oleksandr Tiutyk <trofimich@gmail.com>
SPDX-License-Identifier: MIT
License: https://opensource.org/license/mit
*)

(*!
<summary>Provides fluent assertions on a copied WORD value.</summary>
<description>
Copies actual into persistent instance storage before the entry method returns; literals and expression
results therefore remain valid throughout the immediate chain. Owns no heap allocation or pointed-to resource.
The message prefixes every failure until the next preparation. Finish one chain before starting another on
the owning Assertions provider. Use only from the owning test callback on one task, without reentry.
Obtain this context from the owning provider; direct unprepared use is unsupported.
Expected arguments use the declared IEC type; ordinary compiler conversions happen before comparison.
This context does not depend on another assertion context.
Object metadata is available before preparation; inherited equality compares instance identity.
</description>
*)

{attribute 'no_explicit_call' := 'do not call this function block directly'}
FUNCTION_BLOCK WordAssertionContext EXTENDS TOF_Core.Object
VAR_STAT
	{attribute 'hide'}
	_ClassName : STRING := __POUNAME();
END_VAR
VAR
	_Actual : WORD;
	_TestCase : ITestCase;
	_Message : WSTRING(255);
END_VAR

(*!
<summary>Provides the implementation class name.</summary>
<description>
Borrowed read-only reference to compiler-initialized storage, valid throughout the instance lifetime.
Do not modify the returned reference; no ownership is transferred.
</description>
*)
{attribute 'monitoring' := 'call'}
PROPERTY ClassName : REFERENCE TO STRING
GET
ClassName REF= _ClassName;
END_GET
END_PROPERTY

(*!
<summary>Asserts that the actual value is strictly greater than expected.</summary>
<description>
Records failure without interrupting the callback; preserves the message for the rest of the chain.
</description>
<param name="expected">Expected value converted by the compiler to WORD.</param>
*)
METHOD FINAL IsGreaterThan : REFERENCE TO WordAssertionContext
VAR_INPUT
	expected : WORD;
END_VAR
IF _Actual <= expected THEN
	failComparison(
		expected := expected,
		expectation := "Expected value > "
	);
END_IF

IsGreaterThan REF= THIS^;
END_METHOD

(*!
<summary>Asserts that the actual value meets the inclusive lower boundary.</summary>
<description>
Records failure without interrupting the callback; preserves the message for the rest of the chain.
</description>
<param name="expected">Expected value converted by the compiler to WORD.</param>
*)
METHOD FINAL IsGreaterThanOrEquals : REFERENCE TO WordAssertionContext
VAR_INPUT
	expected : WORD;
END_VAR
IF _Actual < expected THEN
	failComparison(
		expected := expected,
		expectation := "Expected value >= "
	);
END_IF

IsGreaterThanOrEquals REF= THIS^;
END_METHOD

(*!
<summary>Asserts that the actual value is strictly less than expected.</summary>
<description>
Records failure without interrupting the callback; preserves the message for the rest of the chain.
</description>
<param name="expected">Expected value converted by the compiler to WORD.</param>
*)
METHOD FINAL IsLessThan : REFERENCE TO WordAssertionContext
VAR_INPUT
	expected : WORD;
END_VAR
IF _Actual >= expected THEN
	failComparison(
		expected := expected,
		expectation := "Expected value < "
	);
END_IF

IsLessThan REF= THIS^;
END_METHOD

(*!
<summary>Asserts that the actual value meets the inclusive upper boundary.</summary>
<description>
Records failure without interrupting the callback; preserves the message for the rest of the chain.
</description>
<param name="expected">Expected value converted by the compiler to WORD.</param>
*)
METHOD FINAL IsLessThanOrEquals : REFERENCE TO WordAssertionContext
VAR_INPUT
	expected : WORD;
END_VAR
IF _Actual > expected THEN
	failComparison(
		expected := expected,
		expectation := "Expected value <= "
	);
END_IF

IsLessThanOrEquals REF= THIS^;
END_METHOD

(*!
<summary>Provides the library namespace.</summary>
<description>
Borrowed read-only reference to the compiler-initialized namespace, valid throughout the instance lifetime.
Do not modify the returned reference; no ownership is transferred.
</description>
*)
{attribute 'monitoring' := 'call'}
PROPERTY NamespaceName : REFERENCE TO STRING
GET
NamespaceName REF= CurrentNamespace.Name;
END_GET
END_PROPERTY

(*!
<summary>Asserts inequality with the expected value.</summary>
<description>
Records failure without interrupting the callback; preserves the message for the rest of the chain.
</description>
<param name="expected">Expected value converted by the compiler to WORD.</param>
*)
METHOD FINAL NotToBe : REFERENCE TO WordAssertionContext
VAR_INPUT
	expected : WORD;
END_VAR
IF _Actual = expected THEN
	failComparison(
		expected := expected,
		expectation := "Expected value not to be: "
	);
END_IF

NotToBe REF= THIS^;
END_METHOD

(*!
<summary>Copies the actual operand and replaces the chain-wide message.</summary>
<description>
Called by the owning Assertions provider after it verifies the running test case.
No pointer to this method's input storage is retained. The receiver is borrowed until the next preparation;
the owning provider keeps it alive throughout the immediate chain.
</description>
<param name="actual">Value copied into this context.</param>
<param name="testCase">Borrowed failure receiver for the immediate chain.</param>
<param name="message">Copied diagnostic prefix, including empty to clear the previous prefix.</param>
*)
METHOD INTERNAL FINAL Prepare
VAR_INPUT
	actual : WORD;
	testCase : ITestCase;
	message : WSTRING(255);
END_VAR
_Actual := actual;
_TestCase := testCase;
_Message := message;
END_METHOD

(*!
<summary>Reports the byte size of this concrete instance.</summary>
<description>
Includes inline fields and nested instances, but excludes separately allocated payloads.
Obtaining the size does not transfer ownership or validate an arbitrary address.
</description>
*)
{attribute 'monitoring' := 'call'}
PROPERTY SelfSize : ULINT
GET
SelfSize := XSIZEOF(THIS^);
END_GET
END_PROPERTY

(*!
<summary>Asserts equality with the expected value.</summary>
<description>
Records failure without interrupting the callback; preserves the message for the rest of the chain.
</description>
<param name="expected">Expected value converted by the compiler to WORD.</param>
*)
METHOD FINAL ToBe : REFERENCE TO WordAssertionContext
VAR_INPUT
	expected : WORD;
END_VAR
IF _Actual <> expected THEN
	failComparison(
		expected := expected,
		expectation := "Expected: "
	);
END_IF

ToBe REF= THIS^;
END_METHOD

(*!
<summary>Formats a failed typed predicate and reports it with the chain message.</summary>
<description>
Does not change operands or chain state. The receiver retains its first failure. Reporting exceptions
propagate to the enclosing test callback handler; an unprepared receiver is a configuration error.
</description>
<param name="expected">Typed expected operand used only for this diagnostic.</param>
<param name="expectation">Prefix identifying the failed predicate.</param>
*)
METHOD PRIVATE failComparison
VAR_INPUT
	expected : WORD;
	expectation : WSTRING(40);
END_VAR
VAR
	actualText : WSTRING(255);
	expectedText : WSTRING(255);
	diagnostic : TOF_Core.ERROR_MESSAGE;
END_VAR
actualText := TO_WSTRING(TO_UINT(_Actual));
expectedText := TO_WSTRING(TO_UINT(expected));

diagnostic := TOF_Core.WideStrings.Concat255(
	expectation,
	expectedText,
	", but was: ",
	actualText
);

TestServices.ReportAssertionFailure(
	testCase := _TestCase,
	message := _Message,
	sourceClassName := ClassName,
	defaultMessage := diagnostic
);
END_METHOD

END_FUNCTION_BLOCK

// ---- Assertions/TypedContexts/DWordAssertionContext.TcPOU
(*
SPDX-FileCopyrightText: © 2026 Oleksandr Tiutyk <trofimich@gmail.com>
SPDX-License-Identifier: MIT
License: https://opensource.org/license/mit
*)

(*!
<summary>Provides fluent assertions on a copied DWORD value.</summary>
<description>
Copies actual into persistent instance storage before the entry method returns; literals and expression
results therefore remain valid throughout the immediate chain. Owns no heap allocation or pointed-to resource.
The message prefixes every failure until the next preparation. Finish one chain before starting another on
the owning Assertions provider. Use only from the owning test callback on one task, without reentry.
Obtain this context from the owning provider; direct unprepared use is unsupported.
Expected arguments use the declared IEC type; ordinary compiler conversions happen before comparison.
This context does not depend on another assertion context.
Object metadata is available before preparation; inherited equality compares instance identity.
</description>
*)

{attribute 'no_explicit_call' := 'do not call this function block directly'}
FUNCTION_BLOCK DWordAssertionContext EXTENDS TOF_Core.Object
VAR_STAT
	{attribute 'hide'}
	_ClassName : STRING := __POUNAME();
END_VAR
VAR
	_Actual : DWORD;
	_TestCase : ITestCase;
	_Message : WSTRING(255);
END_VAR

(*!
<summary>Provides the implementation class name.</summary>
<description>
Borrowed read-only reference to compiler-initialized storage, valid throughout the instance lifetime.
Do not modify the returned reference; no ownership is transferred.
</description>
*)
{attribute 'monitoring' := 'call'}
PROPERTY ClassName : REFERENCE TO STRING
GET
ClassName REF= _ClassName;
END_GET
END_PROPERTY

(*!
<summary>Asserts that the actual value is strictly greater than expected.</summary>
<description>
Records failure without interrupting the callback; preserves the message for the rest of the chain.
</description>
<param name="expected">Expected value converted by the compiler to DWORD.</param>
*)
METHOD FINAL IsGreaterThan : REFERENCE TO DWordAssertionContext
VAR_INPUT
	expected : DWORD;
END_VAR
IF _Actual <= expected THEN
	failComparison(
		expected := expected,
		expectation := "Expected value > "
	);
END_IF

IsGreaterThan REF= THIS^;
END_METHOD

(*!
<summary>Asserts that the actual value meets the inclusive lower boundary.</summary>
<description>
Records failure without interrupting the callback; preserves the message for the rest of the chain.
</description>
<param name="expected">Expected value converted by the compiler to DWORD.</param>
*)
METHOD FINAL IsGreaterThanOrEquals : REFERENCE TO DWordAssertionContext
VAR_INPUT
	expected : DWORD;
END_VAR
IF _Actual < expected THEN
	failComparison(
		expected := expected,
		expectation := "Expected value >= "
	);
END_IF

IsGreaterThanOrEquals REF= THIS^;
END_METHOD

(*!
<summary>Asserts that the actual value is strictly less than expected.</summary>
<description>
Records failure without interrupting the callback; preserves the message for the rest of the chain.
</description>
<param name="expected">Expected value converted by the compiler to DWORD.</param>
*)
METHOD FINAL IsLessThan : REFERENCE TO DWordAssertionContext
VAR_INPUT
	expected : DWORD;
END_VAR
IF _Actual >= expected THEN
	failComparison(
		expected := expected,
		expectation := "Expected value < "
	);
END_IF

IsLessThan REF= THIS^;
END_METHOD

(*!
<summary>Asserts that the actual value meets the inclusive upper boundary.</summary>
<description>
Records failure without interrupting the callback; preserves the message for the rest of the chain.
</description>
<param name="expected">Expected value converted by the compiler to DWORD.</param>
*)
METHOD FINAL IsLessThanOrEquals : REFERENCE TO DWordAssertionContext
VAR_INPUT
	expected : DWORD;
END_VAR
IF _Actual > expected THEN
	failComparison(
		expected := expected,
		expectation := "Expected value <= "
	);
END_IF

IsLessThanOrEquals REF= THIS^;
END_METHOD

(*!
<summary>Provides the library namespace.</summary>
<description>
Borrowed read-only reference to the compiler-initialized namespace, valid throughout the instance lifetime.
Do not modify the returned reference; no ownership is transferred.
</description>
*)
{attribute 'monitoring' := 'call'}
PROPERTY NamespaceName : REFERENCE TO STRING
GET
NamespaceName REF= CurrentNamespace.Name;
END_GET
END_PROPERTY

(*!
<summary>Asserts inequality with the expected value.</summary>
<description>
Records failure without interrupting the callback; preserves the message for the rest of the chain.
</description>
<param name="expected">Expected value converted by the compiler to DWORD.</param>
*)
METHOD FINAL NotToBe : REFERENCE TO DWordAssertionContext
VAR_INPUT
	expected : DWORD;
END_VAR
IF _Actual = expected THEN
	failComparison(
		expected := expected,
		expectation := "Expected value not to be: "
	);
END_IF

NotToBe REF= THIS^;
END_METHOD

(*!
<summary>Copies the actual operand and replaces the chain-wide message.</summary>
<description>
Called by the owning Assertions provider after it verifies the running test case.
No pointer to this method's input storage is retained. The receiver is borrowed until the next preparation;
the owning provider keeps it alive throughout the immediate chain.
</description>
<param name="actual">Value copied into this context.</param>
<param name="testCase">Borrowed failure receiver for the immediate chain.</param>
<param name="message">Copied diagnostic prefix, including empty to clear the previous prefix.</param>
*)
METHOD INTERNAL FINAL Prepare
VAR_INPUT
	actual : DWORD;
	testCase : ITestCase;
	message : WSTRING(255);
END_VAR
_Actual := actual;
_TestCase := testCase;
_Message := message;
END_METHOD

(*!
<summary>Reports the byte size of this concrete instance.</summary>
<description>
Includes inline fields and nested instances, but excludes separately allocated payloads.
Obtaining the size does not transfer ownership or validate an arbitrary address.
</description>
*)
{attribute 'monitoring' := 'call'}
PROPERTY SelfSize : ULINT
GET
SelfSize := XSIZEOF(THIS^);
END_GET
END_PROPERTY

(*!
<summary>Asserts equality with the expected value.</summary>
<description>
Records failure without interrupting the callback; preserves the message for the rest of the chain.
</description>
<param name="expected">Expected value converted by the compiler to DWORD.</param>
*)
METHOD FINAL ToBe : REFERENCE TO DWordAssertionContext
VAR_INPUT
	expected : DWORD;
END_VAR
IF _Actual <> expected THEN
	failComparison(
		expected := expected,
		expectation := "Expected: "
	);
END_IF

ToBe REF= THIS^;
END_METHOD

(*!
<summary>Formats a failed typed predicate and reports it with the chain message.</summary>
<description>
Does not change operands or chain state. The receiver retains its first failure. Reporting exceptions
propagate to the enclosing test callback handler; an unprepared receiver is a configuration error.
</description>
<param name="expected">Typed expected operand used only for this diagnostic.</param>
<param name="expectation">Prefix identifying the failed predicate.</param>
*)
METHOD PRIVATE failComparison
VAR_INPUT
	expected : DWORD;
	expectation : WSTRING(40);
END_VAR
VAR
	actualText : WSTRING(255);
	expectedText : WSTRING(255);
	diagnostic : TOF_Core.ERROR_MESSAGE;
END_VAR
actualText := TO_WSTRING(TO_UDINT(_Actual));
expectedText := TO_WSTRING(TO_UDINT(expected));

diagnostic := TOF_Core.WideStrings.Concat255(
	expectation,
	expectedText,
	", but was: ",
	actualText
);

TestServices.ReportAssertionFailure(
	testCase := _TestCase,
	message := _Message,
	sourceClassName := ClassName,
	defaultMessage := diagnostic
);
END_METHOD

END_FUNCTION_BLOCK

// ---- Assertions/TypedContexts/LWordAssertionContext.TcPOU
(*
SPDX-FileCopyrightText: © 2026 Oleksandr Tiutyk <trofimich@gmail.com>
SPDX-License-Identifier: MIT
License: https://opensource.org/license/mit
*)

(*!
<summary>Provides fluent assertions on a copied LWORD value.</summary>
<description>
Copies actual into persistent instance storage before the entry method returns; literals and expression
results therefore remain valid throughout the immediate chain. Owns no heap allocation or pointed-to resource.
The message prefixes every failure until the next preparation. Finish one chain before starting another on
the owning Assertions provider. Use only from the owning test callback on one task, without reentry.
Obtain this context from the owning provider; direct unprepared use is unsupported.
Expected arguments use the declared IEC type; ordinary compiler conversions happen before comparison.
This context does not depend on another assertion context.
Object metadata is available before preparation; inherited equality compares instance identity.
</description>
*)

{attribute 'no_explicit_call' := 'do not call this function block directly'}
FUNCTION_BLOCK LWordAssertionContext EXTENDS TOF_Core.Object
VAR_STAT
	{attribute 'hide'}
	_ClassName : STRING := __POUNAME();
END_VAR
VAR
	_Actual : LWORD;
	_TestCase : ITestCase;
	_Message : WSTRING(255);
END_VAR

(*!
<summary>Provides the implementation class name.</summary>
<description>
Borrowed read-only reference to compiler-initialized storage, valid throughout the instance lifetime.
Do not modify the returned reference; no ownership is transferred.
</description>
*)
{attribute 'monitoring' := 'call'}
PROPERTY ClassName : REFERENCE TO STRING
GET
ClassName REF= _ClassName;
END_GET
END_PROPERTY

(*!
<summary>Asserts that the actual value is strictly greater than expected.</summary>
<description>
Records failure without interrupting the callback; preserves the message for the rest of the chain.
</description>
<param name="expected">Expected value converted by the compiler to LWORD.</param>
*)
METHOD FINAL IsGreaterThan : REFERENCE TO LWordAssertionContext
VAR_INPUT
	expected : LWORD;
END_VAR
IF _Actual <= expected THEN
	failComparison(
		expected := expected,
		expectation := "Expected value > "
	);
END_IF

IsGreaterThan REF= THIS^;
END_METHOD

(*!
<summary>Asserts that the actual value meets the inclusive lower boundary.</summary>
<description>
Records failure without interrupting the callback; preserves the message for the rest of the chain.
</description>
<param name="expected">Expected value converted by the compiler to LWORD.</param>
*)
METHOD FINAL IsGreaterThanOrEquals : REFERENCE TO LWordAssertionContext
VAR_INPUT
	expected : LWORD;
END_VAR
IF _Actual < expected THEN
	failComparison(
		expected := expected,
		expectation := "Expected value >= "
	);
END_IF

IsGreaterThanOrEquals REF= THIS^;
END_METHOD

(*!
<summary>Asserts that the actual value is strictly less than expected.</summary>
<description>
Records failure without interrupting the callback; preserves the message for the rest of the chain.
</description>
<param name="expected">Expected value converted by the compiler to LWORD.</param>
*)
METHOD FINAL IsLessThan : REFERENCE TO LWordAssertionContext
VAR_INPUT
	expected : LWORD;
END_VAR
IF _Actual >= expected THEN
	failComparison(
		expected := expected,
		expectation := "Expected value < "
	);
END_IF

IsLessThan REF= THIS^;
END_METHOD

(*!
<summary>Asserts that the actual value meets the inclusive upper boundary.</summary>
<description>
Records failure without interrupting the callback; preserves the message for the rest of the chain.
</description>
<param name="expected">Expected value converted by the compiler to LWORD.</param>
*)
METHOD FINAL IsLessThanOrEquals : REFERENCE TO LWordAssertionContext
VAR_INPUT
	expected : LWORD;
END_VAR
IF _Actual > expected THEN
	failComparison(
		expected := expected,
		expectation := "Expected value <= "
	);
END_IF

IsLessThanOrEquals REF= THIS^;
END_METHOD

(*!
<summary>Provides the library namespace.</summary>
<description>
Borrowed read-only reference to the compiler-initialized namespace, valid throughout the instance lifetime.
Do not modify the returned reference; no ownership is transferred.
</description>
*)
{attribute 'monitoring' := 'call'}
PROPERTY NamespaceName : REFERENCE TO STRING
GET
NamespaceName REF= CurrentNamespace.Name;
END_GET
END_PROPERTY

(*!
<summary>Asserts inequality with the expected value.</summary>
<description>
Records failure without interrupting the callback; preserves the message for the rest of the chain.
</description>
<param name="expected">Expected value converted by the compiler to LWORD.</param>
*)
METHOD FINAL NotToBe : REFERENCE TO LWordAssertionContext
VAR_INPUT
	expected : LWORD;
END_VAR
IF _Actual = expected THEN
	failComparison(
		expected := expected,
		expectation := "Expected value not to be: "
	);
END_IF

NotToBe REF= THIS^;
END_METHOD

(*!
<summary>Copies the actual operand and replaces the chain-wide message.</summary>
<description>
Called by the owning Assertions provider after it verifies the running test case.
No pointer to this method's input storage is retained. The receiver is borrowed until the next preparation;
the owning provider keeps it alive throughout the immediate chain.
</description>
<param name="actual">Value copied into this context.</param>
<param name="testCase">Borrowed failure receiver for the immediate chain.</param>
<param name="message">Copied diagnostic prefix, including empty to clear the previous prefix.</param>
*)
METHOD INTERNAL FINAL Prepare
VAR_INPUT
	actual : LWORD;
	testCase : ITestCase;
	message : WSTRING(255);
END_VAR
_Actual := actual;
_TestCase := testCase;
_Message := message;
END_METHOD

(*!
<summary>Reports the byte size of this concrete instance.</summary>
<description>
Includes inline fields and nested instances, but excludes separately allocated payloads.
Obtaining the size does not transfer ownership or validate an arbitrary address.
</description>
*)
{attribute 'monitoring' := 'call'}
PROPERTY SelfSize : ULINT
GET
SelfSize := XSIZEOF(THIS^);
END_GET
END_PROPERTY

(*!
<summary>Asserts equality with the expected value.</summary>
<description>
Records failure without interrupting the callback; preserves the message for the rest of the chain.
</description>
<param name="expected">Expected value converted by the compiler to LWORD.</param>
*)
METHOD FINAL ToBe : REFERENCE TO LWordAssertionContext
VAR_INPUT
	expected : LWORD;
END_VAR
IF _Actual <> expected THEN
	failComparison(
		expected := expected,
		expectation := "Expected: "
	);
END_IF

ToBe REF= THIS^;
END_METHOD

(*!
<summary>Formats a failed typed predicate and reports it with the chain message.</summary>
<description>
Does not change operands or chain state. The receiver retains its first failure. Reporting exceptions
propagate to the enclosing test callback handler; an unprepared receiver is a configuration error.
</description>
<param name="expected">Typed expected operand used only for this diagnostic.</param>
<param name="expectation">Prefix identifying the failed predicate.</param>
*)
METHOD PRIVATE failComparison
VAR_INPUT
	expected : LWORD;
	expectation : WSTRING(40);
END_VAR
VAR
	actualText : WSTRING(255);
	expectedText : WSTRING(255);
	diagnostic : TOF_Core.ERROR_MESSAGE;
END_VAR
actualText := TO_WSTRING(TO_ULINT(_Actual));
expectedText := TO_WSTRING(TO_ULINT(expected));

diagnostic := TOF_Core.WideStrings.Concat255(
	expectation,
	expectedText,
	", but was: ",
	actualText
);

TestServices.ReportAssertionFailure(
	testCase := _TestCase,
	message := _Message,
	sourceClassName := ClassName,
	defaultMessage := diagnostic
);
END_METHOD

END_FUNCTION_BLOCK

// ---- Assertions/TypedContexts/RealAssertionContext.TcPOU
(*
SPDX-FileCopyrightText: © 2026 Oleksandr Tiutyk <trofimich@gmail.com>
SPDX-License-Identifier: MIT
License: https://opensource.org/license/mit
*)

(*!
<summary>Provides fluent assertions on a copied REAL value.</summary>
<description>
Copies actual into persistent instance storage before the entry method returns; literals and expression
results therefore remain valid throughout the immediate chain. Owns no heap allocation or pointed-to resource.
The message prefixes every failure until the next preparation. Finish one chain before starting another on
the owning Assertions provider. Use only from the owning test callback on one task, without reentry.
Obtain this context from the owning provider; direct unprepared use is unsupported.
Expected arguments use the declared IEC type; ordinary compiler conversions happen before comparison.
This context does not depend on another assertion context.
Object metadata is available before preparation; inherited equality compares instance identity.
Equality and inclusive ordering accept a finite nonnegative LREAL tolerance, default zero. Strict ordering
has no tolerance. Core canonical NaN, infinity and signed-zero rules apply; unequal nonfinite values are
never close. Invalid tolerance records failure without throwing. Tolerance belongs only to that method call.
Inclusive ordering also accepts equality from Core ordering under the target's floating configuration;
exact ToBe and NotToBe still compare canonical bits when tolerance is zero.
</description>
*)

{attribute 'no_explicit_call' := 'do not call this function block directly'}
FUNCTION_BLOCK RealAssertionContext EXTENDS TOF_Core.Object
VAR_STAT
	{attribute 'hide'}
	_ClassName : STRING := __POUNAME();
END_VAR
VAR
	_Actual : REAL;
	_TestCase : ITestCase;
	_Message : WSTRING(255);
END_VAR

(*!
<summary>Provides the implementation class name.</summary>
<description>
Borrowed read-only reference to compiler-initialized storage, valid throughout the instance lifetime.
Do not modify the returned reference; no ownership is transferred.
</description>
*)
{attribute 'monitoring' := 'call'}
PROPERTY ClassName : REFERENCE TO STRING
GET
ClassName REF= _ClassName;
END_GET
END_PROPERTY

(*!
<summary>Asserts that the actual value is strictly greater than expected.</summary>
<description>
Records failure without interrupting the callback; preserves the message for the rest of the chain.
</description>
<param name="expected">Expected value converted by the compiler to REAL.</param>
*)
METHOD FINAL IsGreaterThan : REFERENCE TO RealAssertionContext
VAR_INPUT
	expected : REAL;
END_VAR
VAR
	actualBits : ULINT;
	expectedBits : ULINT;
	comparison : TOF_Core.COMPARISON_RESULT;
END_VAR
actualBits := TestServices.GetCanonicalRealBits(value := _Actual);
expectedBits := TestServices.GetCanonicalRealBits(value := expected);

comparison := TestServices.CompareFloatingValues(
	actualBits := actualBits,
	expectedBits := expectedBits
);

IF comparison <> TOF_Core.COMPARISON_RESULT.FIRST_GREATER_THAN_SECOND THEN
	failComparison(
		expected := expected,
		expectation := "Expected value > "
	);
END_IF

IsGreaterThan REF= THIS^;
END_METHOD

(*!
<summary>Asserts that the actual value meets the inclusive lower boundary.</summary>
<description>
Records failure without interrupting the callback; preserves the message for the rest of the chain.
Uses the canonical floating policy shared by the typed contexts, matching Core semantics, and absolute tolerance.
Invalid tolerance records failure before comparison. The default zero does not affect later assertions in this chain.
</description>
<param name="expected">Expected value converted by the compiler to REAL.</param>
<param name="tolerance">Finite nonnegative absolute distance for this call only; default zero.</param>
*)
METHOD FINAL IsGreaterThanOrEquals : REFERENCE TO RealAssertionContext
VAR_INPUT
	expected : REAL;
	tolerance : LREAL := LREAL#0.0;
END_VAR
VAR
	actualBits : ULINT;
	expectedBits : ULINT;
	comparison : TOF_Core.COMPARISON_RESULT;
	isSatisfied : BOOL;
END_VAR
IF NOT TestServices.IsValidFloatingTolerance(tolerance := tolerance) THEN
	TestServices.ReportAssertionFailure(
		testCase := _TestCase,
		message := _Message,
		sourceClassName := ClassName,
		defaultMessage := "Expected a finite nonnegative comparison tolerance"
	);
	IsGreaterThanOrEquals REF= THIS^;
	RETURN;
END_IF

actualBits := TestServices.GetCanonicalRealBits(value := _Actual);
expectedBits := TestServices.GetCanonicalRealBits(value := expected);

comparison := TestServices.CompareFloatingValues(
	actualBits := actualBits,
	expectedBits := expectedBits
);

isSatisfied := (comparison = TOF_Core.COMPARISON_RESULT.FIRST_GREATER_THAN_SECOND)
	OR_ELSE (comparison = TOF_Core.COMPARISON_RESULT.FIRST_EQUAL_TO_SECOND)
	OR_ELSE TestServices.AreFloatingValuesWithinTolerance(
		actualBits := actualBits,
		expectedBits := expectedBits,
		tolerance := tolerance
	);

IF NOT isSatisfied THEN
	failComparison(
		expected := expected,
		expectation := "Expected value >= ",
		toleranceText := TOF_Core.WideStrings.Concat255(", tolerance: ", TO_WSTRING(tolerance))
	);
END_IF

IsGreaterThanOrEquals REF= THIS^;
END_METHOD

(*!
<summary>Asserts that the actual value is strictly less than expected.</summary>
<description>
Records failure without interrupting the callback; preserves the message for the rest of the chain.
</description>
<param name="expected">Expected value converted by the compiler to REAL.</param>
*)
METHOD FINAL IsLessThan : REFERENCE TO RealAssertionContext
VAR_INPUT
	expected : REAL;
END_VAR
VAR
	actualBits : ULINT;
	expectedBits : ULINT;
	comparison : TOF_Core.COMPARISON_RESULT;
END_VAR
actualBits := TestServices.GetCanonicalRealBits(value := _Actual);
expectedBits := TestServices.GetCanonicalRealBits(value := expected);

comparison := TestServices.CompareFloatingValues(
	actualBits := actualBits,
	expectedBits := expectedBits
);

IF comparison <> TOF_Core.COMPARISON_RESULT.FIRST_LESS_THAN_SECOND THEN
	failComparison(
		expected := expected,
		expectation := "Expected value < "
	);
END_IF

IsLessThan REF= THIS^;
END_METHOD

(*!
<summary>Asserts that the actual value meets the inclusive upper boundary.</summary>
<description>
Records failure without interrupting the callback; preserves the message for the rest of the chain.
Uses the canonical floating policy shared by the typed contexts, matching Core semantics, and absolute tolerance.
Invalid tolerance records failure before comparison. The default zero does not affect later assertions in this chain.
</description>
<param name="expected">Expected value converted by the compiler to REAL.</param>
<param name="tolerance">Finite nonnegative absolute distance for this call only; default zero.</param>
*)
METHOD FINAL IsLessThanOrEquals : REFERENCE TO RealAssertionContext
VAR_INPUT
	expected : REAL;
	tolerance : LREAL := LREAL#0.0;
END_VAR
VAR
	actualBits : ULINT;
	expectedBits : ULINT;
	comparison : TOF_Core.COMPARISON_RESULT;
	isSatisfied : BOOL;
END_VAR
IF NOT TestServices.IsValidFloatingTolerance(tolerance := tolerance) THEN
	TestServices.ReportAssertionFailure(
		testCase := _TestCase,
		message := _Message,
		sourceClassName := ClassName,
		defaultMessage := "Expected a finite nonnegative comparison tolerance"
	);
	IsLessThanOrEquals REF= THIS^;
	RETURN;
END_IF

actualBits := TestServices.GetCanonicalRealBits(value := _Actual);
expectedBits := TestServices.GetCanonicalRealBits(value := expected);

comparison := TestServices.CompareFloatingValues(
	actualBits := actualBits,
	expectedBits := expectedBits
);

isSatisfied := (comparison = TOF_Core.COMPARISON_RESULT.FIRST_LESS_THAN_SECOND)
	OR_ELSE (comparison = TOF_Core.COMPARISON_RESULT.FIRST_EQUAL_TO_SECOND)
	OR_ELSE TestServices.AreFloatingValuesWithinTolerance(
		actualBits := actualBits,
		expectedBits := expectedBits,
		tolerance := tolerance
	);

IF NOT isSatisfied THEN
	failComparison(
		expected := expected,
		expectation := "Expected value <= ",
		toleranceText := TOF_Core.WideStrings.Concat255(", tolerance: ", TO_WSTRING(tolerance))
	);
END_IF

IsLessThanOrEquals REF= THIS^;
END_METHOD

(*!
<summary>Provides the library namespace.</summary>
<description>
Borrowed read-only reference to the compiler-initialized namespace, valid throughout the instance lifetime.
Do not modify the returned reference; no ownership is transferred.
</description>
*)
{attribute 'monitoring' := 'call'}
PROPERTY NamespaceName : REFERENCE TO STRING
GET
NamespaceName REF= CurrentNamespace.Name;
END_GET
END_PROPERTY

(*!
<summary>Asserts inequality with the expected value.</summary>
<description>
Records failure without interrupting the callback; preserves the message for the rest of the chain.
Uses the canonical floating policy shared by the typed contexts, matching Core semantics, and absolute tolerance.
Invalid tolerance records failure before comparison. The default zero does not affect later assertions in this chain.
</description>
<param name="expected">Expected value converted by the compiler to REAL.</param>
<param name="tolerance">Finite nonnegative absolute distance for this call only; default zero.</param>
*)
METHOD FINAL NotToBe : REFERENCE TO RealAssertionContext
VAR_INPUT
	expected : REAL;
	tolerance : LREAL := LREAL#0.0;
END_VAR
VAR
	actualBits : ULINT;
	expectedBits : ULINT;
	areEqual : BOOL;
END_VAR
IF NOT TestServices.IsValidFloatingTolerance(tolerance := tolerance) THEN
	TestServices.ReportAssertionFailure(
		testCase := _TestCase,
		message := _Message,
		sourceClassName := ClassName,
		defaultMessage := "Expected a finite nonnegative comparison tolerance"
	);
	NotToBe REF= THIS^;
	RETURN;
END_IF

actualBits := TestServices.GetCanonicalRealBits(value := _Actual);
expectedBits := TestServices.GetCanonicalRealBits(value := expected);

areEqual := TestServices.AreFloatingValuesWithinTolerance(
	actualBits := actualBits,
	expectedBits := expectedBits,
	tolerance := tolerance
);

IF areEqual THEN
	failComparison(
		expected := expected,
		expectation := "Expected value not to be: ",
		toleranceText := TOF_Core.WideStrings.Concat255(", tolerance: ", TO_WSTRING(tolerance))
	);
END_IF

NotToBe REF= THIS^;
END_METHOD

(*!
<summary>Copies the actual operand and replaces the chain-wide message.</summary>
<description>
Called by the owning Assertions provider after it verifies the running test case.
No pointer to this method's input storage is retained. The receiver is borrowed until the next preparation;
the owning provider keeps it alive throughout the immediate chain.
</description>
<param name="actual">Value copied into this context.</param>
<param name="testCase">Borrowed failure receiver for the immediate chain.</param>
<param name="message">Copied diagnostic prefix, including empty to clear the previous prefix.</param>
*)
METHOD INTERNAL FINAL Prepare
VAR_INPUT
	actual : REAL;
	testCase : ITestCase;
	message : WSTRING(255);
END_VAR
_Actual := actual;
_TestCase := testCase;
_Message := message;
END_METHOD

(*!
<summary>Reports the byte size of this concrete instance.</summary>
<description>
Includes inline fields and nested instances, but excludes separately allocated payloads.
Obtaining the size does not transfer ownership or validate an arbitrary address.
</description>
*)
{attribute 'monitoring' := 'call'}
PROPERTY SelfSize : ULINT
GET
SelfSize := XSIZEOF(THIS^);
END_GET
END_PROPERTY

(*!
<summary>Asserts equality with the expected value.</summary>
<description>
Records failure without interrupting the callback; preserves the message for the rest of the chain.
Uses the canonical floating policy shared by the typed contexts, matching Core semantics, and absolute tolerance.
Invalid tolerance records failure before comparison. The default zero does not affect later assertions in this chain.
</description>
<param name="expected">Expected value converted by the compiler to REAL.</param>
<param name="tolerance">Finite nonnegative absolute distance for this call only; default zero.</param>
*)
METHOD FINAL ToBe : REFERENCE TO RealAssertionContext
VAR_INPUT
	expected : REAL;
	tolerance : LREAL := LREAL#0.0;
END_VAR
VAR
	actualBits : ULINT;
	expectedBits : ULINT;
	areEqual : BOOL;
END_VAR
IF NOT TestServices.IsValidFloatingTolerance(tolerance := tolerance) THEN
	TestServices.ReportAssertionFailure(
		testCase := _TestCase,
		message := _Message,
		sourceClassName := ClassName,
		defaultMessage := "Expected a finite nonnegative comparison tolerance"
	);
	ToBe REF= THIS^;
	RETURN;
END_IF

actualBits := TestServices.GetCanonicalRealBits(value := _Actual);
expectedBits := TestServices.GetCanonicalRealBits(value := expected);

areEqual := TestServices.AreFloatingValuesWithinTolerance(
	actualBits := actualBits,
	expectedBits := expectedBits,
	tolerance := tolerance
);

IF NOT areEqual THEN
	failComparison(
		expected := expected,
		expectation := "Expected: ",
		toleranceText := TOF_Core.WideStrings.Concat255(", tolerance: ", TO_WSTRING(tolerance))
	);
END_IF

ToBe REF= THIS^;
END_METHOD

(*!
<summary>Formats a failed typed predicate and reports it with the chain message.</summary>
<description>
Does not change operands or chain state. The receiver retains its first failure. Reporting exceptions
propagate to the enclosing test callback handler; an unprepared receiver is a configuration error.
</description>
<param name="expected">Typed expected operand used only for this diagnostic.</param>
<param name="expectation">Prefix identifying the failed predicate.</param>
<param name="toleranceText">Optional call-local tolerance suffix; empty for strict ordering.</param>
*)
METHOD PRIVATE failComparison
VAR_INPUT
	expected : REAL;
	expectation : WSTRING(40);
	toleranceText : WSTRING(80) := "";
END_VAR
VAR
	actualText : WSTRING(255);
	expectedText : WSTRING(255);
	diagnostic : TOF_Core.ERROR_MESSAGE;
END_VAR
actualText := TO_WSTRING(_Actual);
expectedText := TO_WSTRING(expected);

